(* IEC 61131-3 sources: codesys-framework/txt/application/WeVe IO (library)/Analog Output, 3 files *)

(* ---- E_AnalogOutputType.dut.st ---- *)
TYPE E_AnalogOutputType :
(
	Invalid := 0,
	S501_0_10V := 1
);
END_TYPE

(* ---- SC_SystemParametersAnalogOutput.dut.st ---- *)
TYPE SC_SystemParametersAnalogOutput :
STRUCT
	eSysPar_AO_Type 								: E_AnalogOutputType;
	eSignalEngUnit 									: E_EngineeringUnits;
	iSysPar_SignalValue_Raw_atAnalogMinLevel 		: INT 	:= 0;
	iSysPar_SignalValue_Raw_atAnalogMaxLevel 		: INT 	:= 16384;
	rSysPar_SignalValue_EngUnit_atAnalogMinLevel 	: REAL;
	rSysPar_SignalValue_EngUnit_atAnalogMaxLevel 	: REAL;
END_STRUCT
END_TYPE

(* ---- FB_AnalogOutput.pou.st ---- *)
FUNCTION_BLOCK FB_AnalogOutput
VAR_INPUT
END_VAR
VAR_OUTPUT
	iAQ_Value 				: INT;
END_VAR
VAR
	_scSysPar 				: SC_SystemParametersAnalogOutput;
	_rSetPoint 				: REAL;
END_VAR

// --- BEGIN IMPLEMENTATION ---

iAQ_Value := REAL_TO_INT (F_Scale (
	rInputScaleValue := _rSetPoint,
	rInputScaleValueMinLevel := _scSysPar.rSysPar_SignalValue_EngUnit_atAnalogMinLevel,
	rInputScaleValueMaxLevel := _scSysPar.rSysPar_SignalValue_EngUnit_atAnalogMaxLevel,
	rOutputScaleValueMinLevel := _scSysPar.iSysPar_SignalValue_Raw_atAnalogMinLevel,
	rOutputScaleValueMaxLevel := _scSysPar.iSysPar_SignalValue_Raw_atAnalogMaxLevel,
	eScaleMethod := E_ScaleMethod.InterPolationZero_whenOutLimits));
